(* IEC 61131-3 sources: SortJet_MasterSPS_Aufbau.fbsproj/Device.device.xml.v3^/Plc Logic.plclogic.xml.v3^/Application.application.xml.v3^/09_Station/Stationen/Kipptisch[206]/0_Konfig, 3 files *)

(* ---- Antriebsinformationen_206.gvl ---- *)
(* METADATA
{
	"v3Meta": {
		"objectGuid": "6a6a4a8e-ada4-4cf2-824b-6c461c89d65a"
	}
}
*)
{attribute 'allow_unqualified_access'}
NAMESPACE Antriebsinformationen_206
VAR_GLOBAL

//-------------------------------------------------------------------------------------------------
// ANTRIEBSINFORMATION [KIPPTISCH]
//-------------------------------------------------------------------------------------------------

  apgInfoStation206Glastransport : ARRAY[cWAND_1..cANZAHL_WAENDE] OF AntriebsInformationen := [
    (
      wAchsID                                 :=      4,  // Achs ID aus dem EConSet
      stTyp                                   := 'Belt',  // Typ
      wpSchaltschrank                         :=   2060,  // Daten aus dem Schaltplan
      wpSchaltplanreihe                       :=     02,  // Daten aus dem Schaltplan
      wpSchaltplanseite                       :=    100,  // Daten aus dem Schaltplan
      rpMaxGeschwindigkeit                    :=   1000,  // [mm/s]   Max- Geschwindigkeit für den Automatikbetrieb
      rpHandGeschwindigkeit                   :=    333,  // [mm/s]   Hand- Geschwindigkeit
      rpReduzierteGeschwindigkeit             :=     67,  // [mm/s]   Reduzierte Geschwindigkeit
      rpReferenzGeschwindigkeit               :=      0,  // [mm/s]   Geschwindigkeit für die Referenzfahrt
      rpEinrichtGeschwindigkeit               :=     50,  // [mm/s]   Max Geschwindigkeit während der Einrichtung der Anlage
      rpMaxBeschleunigung                     :=   1500,  // [mm/s^2] Max Beschleunigung
      rpMaxVerzoegerung                       :=   2000,  // [mm/s^2] Max Verzoegerung
      rpMaxRuckzeit                           :=     50,  // [ms]     Ruckzeit des Antriebs
      rpReduzierteBeschleunigung              :=   1000,  // [mm/s^2] Reduzierte Beschleunigung
      rpReduzierteVerzoegerung                :=   1000,  // [mm/s^2] Reduzierte Verzoegerung
      rpBeschleunigungFremdanlage             :=   1000,  // [mm/s^2] Beschleunigung zu einer Fremdanlage
      rpGeschwindigkeitMessen                 :=    667,  // [mm/s] Geschwindigkeit beim Scheiben messen
      rpGeschwindigkeitSystemcheck            :=  500.0,  // [mm/s]   Geschwindigkeit im Systemcheck (nur Glastransport)
      rpGeschwindigkeitSystemcheckReduzierung :=  167.0,  // [mm/s]   Geschwindigkeit im Systemcheck bei belegtem Vorstop-Sensor (nur Glastransport)
      stOptionen                              := ( eEndschalterQuelle    := Endschalterquelle_EN.KEINE,     // Hardware-Endschalter: KEINE, UMRICHTER oder SPS
                                                   bVersorgungUeberXVR   := FALSE,                          // XVR-Modus: brueckt Hauptschalter 400 V und LS 230 V
                                                   bBremseLoesenFreigabe := FALSE )                         // Der Antrieb darf über eine Betriebsart die Bremse lösen
    )];

  apgInfoStation206Glastransport_Slave : ARRAY[cWAND_1..cANZAHL_WAENDE] OF AntriebsInformationen := [
    (
      wAchsID                                 :=     5,   // Achs ID aus dem EConSet
      stTyp                                   := 'Rolls', // Typ
      wpSchaltschrank                         :=   2061,  // Daten aus dem Schaltplan
      wpSchaltplanreihe                       :=     02,  // Daten aus dem Schaltplan
      wpSchaltplanseite                       :=    100,  // Daten aus dem Schaltplan
      rpMaxGeschwindigkeit                    :=   1000,  // [mm/s]   Max- Geschwindigkeit für den Automatikbetrieb
      rpHandGeschwindigkeit                   :=    333,  // [mm/s]   Hand- Geschwindigkeit
      rpReduzierteGeschwindigkeit             :=     67,  // [mm/s]   Reduzierte Geschwindigkeit
      rpReferenzGeschwindigkeit               :=      0,  // [mm/s]   Geschwindigkeit für die Referenzfahrt
      rpEinrichtGeschwindigkeit               :=     50,  // [mm/s]   Max Geschwindigkeit während der Einrichtung der Anlage
      rpMaxBeschleunigung                     :=   1500,  // [mm/s^2] Max Beschleunigung
      rpMaxVerzoegerung                       :=   2000,  // [mm/s^2] Max Verzoegerung
      rpMaxRuckzeit                           :=     50,  // [ms]     Ruckzeit des Antriebs
      rpReduzierteBeschleunigung              :=   1000,  // [mm/s^2] Reduzierte Beschleunigung
      rpReduzierteVerzoegerung                :=   1000,  // [mm/s^2] Reduzierte Verzoegerung
      rpBeschleunigungFremdanlage             :=   1000,  // [mm/s^2] Beschleunigung zu einer Fremdanlage
      rpGeschwindigkeitMessen                 :=    667,  // [mm/s] Geschwindigkeit beim Scheiben messen
      rpGeschwindigkeitSystemcheck            :=  500.0,  // [mm/s]   Geschwindigkeit im Systemcheck (nur Glastransport)
      rpGeschwindigkeitSystemcheckReduzierung :=  167.0,  // [mm/s]   Geschwindigkeit im Systemcheck bei belegtem Vorstop-Sensor (nur Glastransport)
      stOptionen                              := ( eEndschalterQuelle    := Endschalterquelle_EN.KEINE,     // Hardware-Endschalter: KEINE, UMRICHTER oder SPS
                                                   bVersorgungUeberXVR   := FALSE,                          // XVR-Modus: brueckt Hauptschalter 400 V und LS 230 V
                                                   bBremseLoesenFreigabe := FALSE )                         // Der Antrieb darf über eine Betriebsart die Bremse lösen
    )];

  apgInfoStation206Kippen : AntriebsInformationen :=
    (
      wAchsID                                 :=      6,  // Achs ID aus dem EConSet
      stTyp                                   := 'Tilt',  // Typ
      wpSchaltschrank                         :=   2062,  // Daten aus dem Schaltplan
      wpSchaltplanreihe                       :=      2,  // Daten aus dem Schaltplan
      wpSchaltplanseite                       :=    100,  // Daten aus dem Schaltplan
      rpMaxGeschwindigkeit                    :=     90,  // [Grad/s]   Max- Geschwindigkeit für den Automatikbetrieb // 103 MAX
      rpHandGeschwindigkeit                   :=     40,  // [Grad/s]   Hand- Geschwindigkeit
      rpReduzierteGeschwindigkeit             :=     60,  // [Grad/s]   Reduzierte Geschwindigkeit
      rpReferenzGeschwindigkeit               :=      2,  // [Grad/s]   Geschwindigkeit für die Referenzfahrt
      rpEinrichtGeschwindigkeit               :=      1,  // [Grad/s]   Max Geschwindigkeit während der Einrichtung der Anlage
      rpMaxBeschleunigung                     :=    500,  // [Grad/s^2] Max Beschleunigung
      rpMaxVerzoegerung                       :=    500,  // [Grad/s^2] Max Verzoegerung
      rpMaxRuckzeit                           :=    500,  // [ms] Ruckzeit des Antriebs
      rpReduzierteBeschleunigung              :=    100,  // [Grad/s^2] Reduzierte Beschleunigung
      rpReduzierteVerzoegerung                :=     50,  // [Grad/s^2] Reduzierte Verzoegerung
      rpBeschleunigungFremdanlage             :=      2,  // [Grad/s^2] Beschleunigung zu einer Fremdanlage
      rpGeschwindigkeitMessen                 := 0.0,  // [Grad/s] Geschwindigkeit für die Messfahrt
      rpGeschwindigkeitSystemcheck            :=  500.0,  // [mm/s]   Geschwindigkeit im Systemcheck (nur Glastransport)
      rpGeschwindigkeitSystemcheckReduzierung :=  167.0,  // [mm/s]   Geschwindigkeit im Systemcheck bei belegtem Vorstop-Sensor (nur Glastransport)
      stOptionen                              := ( eEndschalterQuelle    := Endschalterquelle_EN.UMRICHTER, // Hardware-Endschalter: KEINE, UMRICHTER oder SPS
                                                   bVersorgungUeberXVR   := FALSE,                          // XVR-Modus: brueckt Hauptschalter 400 V und LS 230 V
                                                   bBremseLoesenFreigabe := FALSE )                         // Der Antrieb darf über eine Betriebsart die Bremse lösen
    );

  // Querfahrt
  apgInfoStation206Querfahrt : AntriebsInformationen :=
    (
      wAchsID                                 :=        65,  // Achs ID aus dem EConSet
      stTyp                                   := 'Lateral',  // Typ
      wpSchaltschrank                         :=      2063,  // Daten aus dem Schaltplan
      wpSchaltplanreihe                       :=        02,  // Daten aus dem Schaltplan
      wpSchaltplanseite                       :=         0,  // Daten aus dem Schaltplan
      rpMaxGeschwindigkeit                    :=      1000,  // [mm/s]   Max- Geschwindigkeit für den Automatikbetrieb
      rpHandGeschwindigkeit                   :=      1000,  // [mm/s]   Hand- Geschwindigkeit
      rpReduzierteGeschwindigkeit             :=        25,  // [mm/s]   Reduzierte Geschwindigkeit
      rpReferenzGeschwindigkeit               :=        10,  // [mm/s]   Geschwindigkeit für die Referenzfahrt
      rpEinrichtGeschwindigkeit               :=        10,  // [mm/s]   Max Geschwindigkeit während der Einrichtung der Anlage
      rpMaxBeschleunigung                     :=       500,  // [mm/s^2] Max Beschleunigung
      rpMaxVerzoegerung                       :=       500,  // [mm/s^2] Max Verzoegerung
      rpMaxRuckzeit                           :=      1000,  // [ms]     Ruckzeit des Antriebs
      rpReduzierteBeschleunigung              :=        10,  // [mm/s^2] Reduzierte Beschleunigung
      rpReduzierteVerzoegerung                :=        10,  // [mm/s^2] Reduzierte Verzoegerung
      rpBeschleunigungFremdanlage             :=         0,  // [mm/s^2] Beschleunigung zu einer Fremdanlage
      rpGeschwindigkeitMessen                 :=         0,  // [mm/s] Geschwindigkeit beim Scheiben messen
      rpGeschwindigkeitSystemcheck            :=     500.0,  // [mm/s]   Geschwindigkeit im Systemcheck (nur Glastransport)
      rpGeschwindigkeitSystemcheckReduzierung :=     167.0,  // [mm/s]   Geschwindigkeit im Systemcheck bei belegtem Vorstop-Sensor (nur Glastransport)
      stOptionen                              := ( eEndschalterQuelle    := Endschalterquelle_EN.UMRICHTER, // Hardware-Endschalter: KEINE, UMRICHTER oder SPS
                                                   bVersorgungUeberXVR   := FALSE,                          // XVR-Modus: brueckt Hauptschalter 400 V und LS 230 V
                                                   bBremseLoesenFreigabe := FALSE )                         // Der Antrieb darf über eine Betriebsart die Bremse lösen
    );

END_VAR

END_NAMESPACE

(* ---- MK_Station_206.gvl ---- *)
(* METADATA
{
	"v3Meta": {
		"objectGuid": "d056a025-7346-4412-a27e-a3ba4851b2d6"
	}
}
*)
{attribute 'allow_unqualified_access'}
NAMESPACE MK_Station_206
VAR_GLOBAL

//-------------------------------------------------------------------------------------------------
// MASCHINEPARAMETER: KIPPTISCH
//-------------------------------------------------------------------------------------------------

  apgMKStation206 : Parameter_Station:=
    (
      stStationsNummern                     := ( NummerIntern :=   206,                                                    // Stationsnummer fuer das MMI und die Stationsangabe der Meldungen
                                                 NummerExtern :=  1206,                                                    // Stationsnummer fuer Bedienermeldungen
                                                 NummerSPS    :=   206 ),                                                  // Stationsnummer SPS-intern (Indizes)
      bDeaktivieren                         := FALSE,                                                                      // Station deaktiviert (keine Auftraege, keine Referenzfahrt)
      wMeldungsNummer                       := 1790,                                                                       // Basis-Meldungsnummer (WatchIO)
      eStationsTyp                          := eStation,                                                                   // Typ der Station
      eaAutomatikkreis                      := [eAutomatikkreis_1],                                                        // Automatikkreise, zu denen die Station gehoert
      eaSicherheitskreis                    := [eSicherheitskreis_1],                                                      // Sicherheitskreise, in die die Station eingebunden ist
      // astSicherheitskreisTeilabschaltung
      eSystemcheckZyklus                    := eSystemcheckZyklus_1,                                                       // In welchem Zyklus des Systemchecks die Station geprueft wird
      stSchnittstellendaten                 := ( wVorgaengerStation := cSTATION_204,                                       // Station vor dieser Station (cSTATION_DYNAMISCH bei mehreren)
                                                 wNachfolgerStation := cSTATION_207,                                       // Station nach dieser Station (cSTATION_DYNAMISCH bei mehreren)
                                                 bStationIstShuttle := FALSE                                               // Station ist ein Shuttle
                                               ),
      stStationsOptionen                    := ( stSystemcheck :=  ( bScheibenVermessenSystemCheck               := TRUE,  // Scheiben im Systemcheck vermessen
                                                                     bScheibeNachSystemcheckAufAuslauf           := TRUE,  // Scheibe nach dem Systemcheck auf den Auslaufsensor fahren
                                                                     bSystemCheckMitVorgaengerBatchTransport     := FALSE, // derzeit ohne Funktion
                                                                     bSystemCheckMitNachfolgerBatchTransport     := FALSE, // derzeit ohne Funktion
                                                                     bOptionSystemCheckScheibeMittigLegen        := FALSE  // derzeit ohne Funktion
                                                                    ),

                                                 // stTransfershuttle
                                                 stGlastransport :=  ( bVortransport                             := FALSE, // Vortransport aktivieren [Bsp.: Nach einem Eintransport mit gesetztem Bit <Letzte Scheibe>]
                                                                       bTransportMasterSlaveEintransport         := FALSE, // derzeit ohne Funktion
                                                                       bTransportMasterSlaveAustransport         := TRUE , // Austransport als Slave auf die Achse des Nachfolgers
                                                                       bGLasUebernahmeSenkrecht                  := FALSE, // RKT - Eintransport in Senkrechter-Position bzw. in Waagerechter- Position [default]
                                                                       bAustransportISOLinie                     := FALSE, // Austransport an eine ISO-Linie
                                                                       bScheibenVermessen                        := FALSE, // Scheibenmessung am Anlegetisch/Anlegewand
                                                                       bMessrichtungNegativ                      := FALSE, // Negative Fahrtrichtung beim Messen
                                                                       bScheibenmessungEintransport              := FALSE, // Scheibenmessung beim Eintransport
                                                                       bScheibenmessungSensorVorabAuslauf        := FALSE  // Scheibenmessung mit SensorVorabAuslauf z.B. Anlegewand
                                                                      ),
                                                 // stAnlegetisch
                                                 // stEckuebergabe
                                                 // stDrehstation
                                                 bVorAbKomponentenAnsteuerung              := FALSE,                       // VorAbKomponentenAnsteuerung Auftraege werden bearbeitet
                                                 bVerstellungEinAusGefahrenLogikDrehen     := FALSE,                       // Verstellung: Logik ein-/ausgefahren gedreht
                                                 bLangsamfahrtNockenQuerfahrtAktivieren    := FALSE,                       // Querfahrt: Langsamfahrt-Nocken auswerten
                                                 bSKBlockierenDurchVorabSensoren           := FALSE,                       // Vorab-Sensoren belegt blockieren das Oeffnen des Sicherheitskreises
                                                 bStationLeerfahrenBeiSkAnforderung        := FALSE,                       // Station bei Anforderung Sicherheitskreis leerfahren
                                                 bGlasAbgenommenAutomatischQuittieren      := FALSE,                       // derzeit ohne Funktion
                                                 bScheibeAbnehmenNachEintransport          := FALSE                        // Scheibe nach dem Eintransport wieder abnehmen
                                               ),
      stStationsAufbau                      := ( bGeblase                      := [ cANZAHL_WAENDE(FALSE) ],               // Ausbaustufe: Geblaese je Wand
                                                 bGlastransport                := [ TRUE ],                                // Ausbaustufe: Glastransport je Wand
                                                 bKippen                       := [ TRUE ],                                // Ausbaustufe: Kippen je Wand
                                                 bKippenSchuetz                := FALSE,                                   // Kippen ueber Schuetz statt Umrichter
                                                 bTransportVerstellung         := [ cANZAHL_WAENDE(FALSE) ],               // Ausbaustufe Shuttle: Transport-/Dickenverstellung je Wand
                                                 bHub                          := FALSE,                                   // Ausbaustufe: Hub der Station
                                                 bHubrahmen                    := FALSE,                                   // Ausbaustufe: Hubrahmen (Riemen heben/senken)
                                                 bDrehen                       := FALSE,                                   // Ausbaustufe: Drehen
                                                 bQuerachse                    := FALSE,                                   // Ausbaustufe: Querachse
                                                 bMessachse                    := FALSE,                                   // Ausbaustufe: Messachse (Anlegetisch, Anlegewand)
                                                 bDruckluft                    := FALSE,                                   // Druckluftueberwachung vorhanden
                                                 bAnschlag                     := FALSE,                                   // Ausbaustufe: Ausrichtanschlaege
                                                 bSensorAuslauf                := TRUE,                                    // Auslaufsensor vorhanden
                                                 bSensorEinlauf                := TRUE,                                    // Einlaufsensor vorhanden
                                                 bSensorEinlaufStopp           := FALSE,                                   // Shuttle: zusaetzlicher Stopp-Sensor am Einlauf (ohne: Einlaufsensor), Gegenstueck zum Auslauf-Stopp im Rueckwaertstransport
                                                 bSensorAuslaufStopp           := FALSE,                                   // Shuttle: zusaetzlicher Stopp-Sensor am Auslauf (ohne: Auslaufsensor), Verfahrfreigabe und Scheibe hat Shuttle verlassen
                                                 bDurchlaufSperreZumNachfolger := FALSE,                                   // Ausbaustufe: bewegliche Abschrankung zum Nachfolger
                                                 bQuerfahrt                    := FALSE,                                   // Ausbaustufe: Querfahrt
                                                 bKipparme                     := FALSE,                                   // Ausbaustufe: Kipparme
                                                 bSlaveAntrieb                 := TRUE,                                    // Glastransport mit Slave-Antrieb
                                                 bMessachseAmEndeVomTisch      := FALSE,                                   // Messachse am Ende des Tisches (Hoehenfehler fragt den Bediener)
                                                 bWandverstellung              := [ FALSE ],                               // Ausbaustufe Station: Wandverstellung je Wand
                                                 bWandverstellungMotorisch     := FALSE,                                   // Shuttle: Transport-/Wandverstellung mit Antrieb statt pneumatisch
                                                 bRoellchenleiste              := [ FALSE ],                               // Ausbaustufe Station: Roellchenleiste je Wand
                                                 bDurchgang                    := FALSE,                                   // Station ist Teil eines Durchgangs (belegt = Oeffnen blockiert)
                                                 bRolltor                      := FALSE,                                   // Ausbaustufe Faecherwagen: Rolltor
                                                 bKlemmzylinder                := FALSE,                                   // Ausbaustufe Faecherwagen: Klemmzylinder fixiert den Oberrahmen beim Ein- und Ausschleusen
                                                 bGreifer                      := [cANZAHL_WAENDE(FALSE)],                 // Shuttle: Greifer je Wand (Scheibe aus dem Faecherwagen ziehen bzw. hineinschieben)
                                                 bRFID                         := FALSE,                                   // RFID-Leser vorhanden
                                                 bAGV                          := FALSE,                                   // Ausbaustufe Faecherwagen: Betrieb mit AGV
                                                 bDLSSchmiersystem             := FALSE,                                   // Zentralschmierung DLS vorhanden
                                                 bGlastransportSlaveVorhanden  := FALSE,                                   // Glastransport mit Slave-Antrieb (Meldungen/Ueberwachung Slave)
                                                 wHydraulikstation             := 0                                        // Faecherwagen Hydraulik: zugeordnete Hydraulikstation (cHYDRAULIKSTATION_x), 0 = keine
                                               ),
      stStationsParameter                   := ( rLaengeUebergroesseScheibe              := 4240,                          // Shuttle: ab dieser Scheibenlaenge gilt die Scheibe als uebergross [mm]
                                                 rMinGlasHoeheAutomatischenEintransport  := 500,                           // VSG: Mindesthoehe fuer automatischen Eintransport [mm]
                                                 rMinGlasLaengeAutomatischenEintransport := 500,                           // VSG: Mindestlaenge fuer automatischen Eintransport [mm]
                                                 wMaximaleAnzahlAktiverAuftraege := 1,                                     // derzeit ohne Funktion
                                                 rMinPosSwEsEingrenzung                  := 0.0,                           // Externer zusaetzlicher Software-Endschalter MIN; 0 = inaktiv; darf den MK-MIN nur weiter eingrenzen
                                                 rMaxPosSwEsEingrenzung                  := 0.0,                           // Externer zusaetzlicher Software-Endschalter MAX; 0 = inaktiv; darf den MK-MAX nur weiter eingrenzen
                                                 rPosFreigabePufferAusfahren             := 0.0                            // derzeit ohne Funktion
                                              ),
      // stFremdanlage
      stGlasdaten                           := [( rlMinGlasLaenge := 350,                                                  // minimal zulässige GlasLänge
                                                  rlMaxGlasLaenge := 2500,                                                 // maximale zulässige GlasLänge
                                                  rlMinGlasHoehe  := 190,                                                  // minimal zulässige GlasHöhe
                                                  rlMaxGlasHoehe  := 1800,                                                 // maximale zulässige GlasHöhe
                                                  rlMinGlasDicke  := 3,                                                  // minimal zulässige GlasDicke
                                                  rlMaxGlasDicke  := 12.76,                                                   // maximal zulaessige Glasdicke [mm]
                                                  rlLaengeMaxGlas := 0.0                                                   // maximal zulaessige Glaslaenge [mm]
                                               )]
      // astShuttleAnhaltenQuellen
     );

  apgMKStation206Glastransport : ARRAY[cWAND_1..cANZAHL_WAENDE] OF Parameter_Glastransport := [
    (
      rLaengeStation                        := 4800, // Länge der Station
      rScheibenabstand                      :=  300, // Der Abstand zwischen zwei Scheiben auf der Station
      rWegUeberAuslauf                      :=   50, // Weg ueber den Auslaufsensor hinaus [mm]
      rWegUeberEinlauf                      :=   50, // Weg ueber den Einlaufsensor hinaus [mm]
      rWegUeberSensorenSystemCheck          :=   15, // Der Weg der Ueber ein die Sensoren zum vermessen der Scheiben
      rUeberwachungAuslaufsensor            :=  500, // Ueberwachung des Auslaufsensors [Strecke in der der Auslaufsensor Frei / ueberfahren werden soll]
      rUeberwachungEinlaufsensor            :=  500, // Ueberwachung des Einlaufsensors [Strecke in der der Einlaufsensor Frei / ueberfahren werden soll]
      rWegUeberEinlaufEintransport          :=  150, // Eintransport vorwaerts: Abstand Scheibenhinterkante zum Einlaufsensor [mm]
      rWegUeberEinlaufAustransport          :=   50, // Lage Auf Einlauf: Scheibe liegt um diesen Weg auf dem Einlaufsensor [mm]
      rWegUeberAuslaufEintransport          :=   50, // Eintransport rueckwaerts: Abstand Scheibenhinterkante zum Auslaufsensor [mm]
      rWegUeberAuslaufAustransport          :=   50, // Lage Auf Auslauf: Weg ueber den Auslaufsensor hinaus [mm]
      rWegEinlaufsensorZuVorStopSensor      := 4700, // Beschreibt den Weg vum eine Scheibe beim EIntransport vom Einlaufsensor bis ueberden Vorabstopsensor zu verfahren
      rMesstoleranz                         :=   10, // Toleranz-Mass fuer die Scheibenlaengenmessung
      rMessstrecke                          := 4755, // Beschreibt die Strecke ziwischen 2 Sensoren die der Antrieb verfaehrt
      rWegstreckeBisZurVerzoegerung         := 4200  // Beschreibt die Strecke die gefahren werden soll bis der Antrieb abgebremst werden soll, dies gilt fuer Eintransportauftraege die das Bit "Letzte Scheibe" gesetzt haben
    )];

  apgMKStation206Querfahrt : Parameter_Querfahrt :=
    (
      tZeitAntriebsfreigabeErhalten          := T#3M // Energieeinsparung: Zeit nach der die Antriebsfreigabe entzogen wird, wenn keine Aktion ansteht
    );

  apgMKStation206Kippen : ARRAY[cWAND_1..cANZAHL_WAENDE] OF Parameter_Kippen := [
    (
      tZeitlicheUeberwachungKippen          := TIME#5000MS, // [ms \ s] Verwendet fuer Antriebe die Ueber einen Schuetz angesteuert werden
      tZeitAntriebsfreigabeErhalten         :=   TIME#180S, // [ms \ s] Energieeinsparrung: Zeiteinheit nach der die Antriebsfreigabe entzogen werden soll wenn keine Aktion ansteht [1 s = 1000 ms ]
      rToleranz                             :=           1, // Toleranz beim Entscheiden der aktuellen Position
      rPosition0Grad                        :=           0, // Waagerechte- Position 0 Grad: Position auf die die Station gehoben werden soll
      rPosition84Grad                       :=      224.64, // Senkrechte- Position 84 Grad: Position auf die die Station gehoben werden soll
      rPosition90Grad                       :=      224.64, // Senkrechte-Position 90 Grad : Position auf die die Station gesenkt werden soll
      bKippenMitSchuetz                     :=       FALSE, // Kippen per Umrichter oder Schütz
      rPosition88_5Grad                     := 0.0,         // Senkrechte- Position 84 Grad: Position auf die die Station gehoben werden soll
      rPosition96Grad                       := 0.0          // Senkrechte-Position 96 Grad : Position auf die die Station gesenkt werden soll
    )];

END_VAR
END_NAMESPACE

(* ---- Konfiguration_206.gvl ---- *)
(* METADATA
{
	"v3Meta": {
		"objectGuid": "42ae5482-243e-48a3-a681-16c36dcef6f3"
	}
}
*)
{attribute 'allow_unqualified_access'}
NAMESPACE Konfiguration_206
VAR_CONFIG
//-------------------------------------------------------------------------------------------------
// KONFIGURATION: BAUSTEIN IO´s
//-------------------------------------------------------------------------------------------------

  // Rollenleiste (Zylinder 1: Geoeffnet = ausgefahren, Geschlossen = eingefahren; Zylinder 2 ohne Funktion)
  Globale_Bausteine.Kipptisch206.Rollenleiste.in_bStatusZylinder1Ausgefahren                      AT %MX1.0   : BOOL; // OPTION
  Globale_Bausteine.Kipptisch206.Rollenleiste.in_bStatusZylinder1Eingefahren                      AT %MX1.0   : BOOL; // OPTION
  Globale_Bausteine.Kipptisch206.Rollenleiste.in_bStatusZylinder2Ausgefahren                      AT %MX1.0   : BOOL; // OPTION
  Globale_Bausteine.Kipptisch206.Rollenleiste.in_bStatusZylinder2Eingefahren                      AT %MX1.0   : BOOL; // OPTION
  Globale_Bausteine.Kipptisch206.Rollenleiste.out_bZylinder1Ausfahren                             AT %MX2060.0 : BOOL; // OPTION
  Globale_Bausteine.Kipptisch206.Rollenleiste.out_bZylinder1Einfahren                             AT %MX2060.1 : BOOL; // OPTION
  Globale_Bausteine.Kipptisch206.Rollenleiste.out_bZylinder2Ausfahren                             AT %MX2060.2 : BOOL; // OPTION
  Globale_Bausteine.Kipptisch206.Rollenleiste.out_bZylinder2Einfahren                             AT %MX2060.3 : BOOL; // OPTION

  // Kippen
  Globale_Bausteine.Kipptisch206.Kippen.in_bMotorstarter_OK                                       AT %MX1.1   : BOOL; // OPTION
  Globale_Bausteine.Kipptisch206.Kippen.in_bLS400V_OK                                             AT %MX1.1   : BOOL; // OPTION
  Globale_Bausteine.Kipptisch206.Kippen.in_bLSBremse_OK                                           AT %MX1.1   : BOOL; // OPTION
  Globale_Bausteine.Kipptisch206.Kippen.out_bKippen84Grad                                         AT %MX2060.4 : BOOL; // OPTION
  Globale_Bausteine.Kipptisch206.Kippen.out_bKippen90Grad                                         AT %MX2060.5 : BOOL; // OPTION
  Globale_Bausteine.Kipptisch206.Kippen.out_bBremseLoesen                                         AT %MX2060.6 : BOOL; // OPTION
  Globale_Bausteine.Kipptisch206.Kippen.out_bReset                                                AT %MX2060.7 : BOOL; // OPTION

  // Hub (unbenutzt)
  Globale_Bausteine.Kipptisch206.HubUnbenutzt.in_bSensorNichtUnten                                AT %MX1.0   : BOOL; // OPTION
  Globale_Bausteine.Kipptisch206.HubUnbenutzt.in_bSensorNichtOben                                 AT %MX1.0   : BOOL; // OPTION
  Globale_Bausteine.Kipptisch206.HubUnbenutzt.in_bMotorstarter_OK                                 AT %MX1.1   : BOOL; // OPTION
  Globale_Bausteine.Kipptisch206.HubUnbenutzt.in_bLSBremse_OK                                     AT %MX1.1   : BOOL; // OPTION
  Globale_Bausteine.Kipptisch206.HubUnbenutzt.in_bLS400V_OK                                       AT %MX1.1   : BOOL; // OPTION
  Globale_Bausteine.Kipptisch206.HubUnbenutzt.out_bHubAbSetzen                                    AT %MX2061.0 : BOOL; // OPTION
  Globale_Bausteine.Kipptisch206.HubUnbenutzt.out_bHubAufSetzen                                   AT %MX2061.1 : BOOL; // OPTION
  Globale_Bausteine.Kipptisch206.HubUnbenutzt.out_bReset                                          AT %MX2061.2 : BOOL; // OPTION
  Globale_Bausteine.Kipptisch206.HubUnbenutzt.out_bBremseLoesen                                   AT %MX2061.3 : BOOL; // OPTION

  // Wandverstellung (unbenutzt)
  Globale_Bausteine.Kipptisch206.WandverstellungUnbenutzt.in_bStatusZylinder1Ausgefahren          AT %MX1.0   : BOOL; // OPTION
  Globale_Bausteine.Kipptisch206.WandverstellungUnbenutzt.in_bStatusZylinder1Eingefahren          AT %MX1.0   : BOOL; // OPTION
  Globale_Bausteine.Kipptisch206.WandverstellungUnbenutzt.in_bStatusZylinder2Ausgefahren          AT %MX1.0   : BOOL; // OPTION
  Globale_Bausteine.Kipptisch206.WandverstellungUnbenutzt.in_bStatusZylinder2Eingefahren          AT %MX1.0   : BOOL; // OPTION
  Globale_Bausteine.Kipptisch206.WandverstellungUnbenutzt.out_bZylinder1Ausfahren                 AT %MX2061.4 : BOOL; // OPTION
  Globale_Bausteine.Kipptisch206.WandverstellungUnbenutzt.out_bZylinder1Einfahren                 AT %MX2061.5 : BOOL; // OPTION
  Globale_Bausteine.Kipptisch206.WandverstellungUnbenutzt.out_bZylinder2Ausfahren                 AT %MX2061.6 : BOOL; // OPTION
  Globale_Bausteine.Kipptisch206.WandverstellungUnbenutzt.out_bZylinder2Einfahren                 AT %MX2061.7 : BOOL; // OPTION

  // Geblaese-Baustein (unbenutzt)
  Globale_Bausteine.Kipptisch206.GeblaeseUnbenutzt.in_bMotorschutzschalter_OK                     AT %MX1.1   : BOOL; // OPTION
  Globale_Bausteine.Kipptisch206.GeblaeseUnbenutzt.out_bStarteGeblaese                            AT %MX2062.0 : BOOL; // OPTION

END_VAR

END_NAMESPACE
